// TIA Portal V19 export
// export: Created 2026-10-15T09:44:24.5896701Z, ExportSetting WithDefaults, DisplayName Totally Integrated Automation Portal, DisplayVersion V19, DisplayName TIA Portal Openness, DisplayVersion V19, DisplayName TIA Portal Version Control Interface, DisplayVersion V19, DisplayName STEP 7 Professional, DisplayVersion V19, DisplayName STEP 7 Safety, DisplayVersion V19, DisplayName WinCC Basic/Comfort/Advanced, DisplayVersion V19, DisplayName WinCC Unified, DisplayVersion V19
FUNCTION "ROLL_PB19" : Void   // FC27, SCL
{ S7_Optimized_Access := 'TRUE' }
VERSION : 0.1
// stored: AutoNumber true, IsIECCheckEnabled false, SetENOAutomatically false, UDAEnableTagReadback false
   VAR_TEMP
      r : Bool;
      a1 : Word;
      a2 : Word;
      activeDataBlock : Int;
      comparisonResults : Array[0..0] of Bool;
   END_VAR
BEGIN

   #r := FALSE;
   #a1 := W#16#0000;
   #a2 := W#16#0000;
   #activeDataBlock := 0;
   // PB19, STEP 5 network 1
   #r := ((NOT "ROLL_IO".Input[3, 6]) AND (NOT "ROLL_State".M[5, 6]) AND (NOT "ROLL_State".M[6, 0]) AND (NOT "ROLL_State".M[6, 2]) AND ("ROLL_IO".Input[3, 1] OR "ROLL_State".M[31, 5]) AND "ROLL_IO".Input[5, 2] AND "ROLL_IO".Input[5, 4] AND "ROLL_State".M[4, 1]);
   "ROLL_State".M[82, 0] := #r;
   // PB19, STEP 5 network 2
   #r := ((NOT "ROLL_IO".Input[3, 6]) AND (NOT "ROLL_State".M[12, 0]) AND (NOT "ROLL_State".M[5, 3]) AND (NOT "ROLL_State".M[5, 6]) AND ("ROLL_IO".Input[3, 1] OR "ROLL_State".M[31, 5]) AND "ROLL_IO".Input[8, 3] AND "ROLL_IO".Input[8, 5] AND "ROLL_State".M[4, 1]);
   "ROLL_State".M[82, 2] := #r;
   // PB19, STEP 5 network 3
   #r := ("ROLL_State".M[31, 5] AND "ROLL_State".M[40, 0]);
   IF #r THEN
       "ROLL_State".M[82, 3] := TRUE;
   END_IF;
   #r := (NOT "ROLL_State".M[31, 5]);
   IF #r THEN
       "ROLL_State".M[82, 3] := FALSE;
   END_IF;
   // PB19, STEP 5 network 4
   #r := ((NOT "ROLL_State".M[110, 1]) AND (NOT "ROLL_State".M[110, 2]) AND "ROLL_State".M[110, 0] AND "ROLL_State".M[110, 3] AND "ROLL_State".M[40, 0]);
   "ROLL_State".M[240, 0] := #r;
   // PB19, STEP 5 network 5
   #r := (((NOT "ROLL_State".M[110, 2]) AND "ROLL_State".M[110, 0] AND "ROLL_State".M[110, 1] AND "ROLL_State".M[110, 3] AND "ROLL_State".M[41, 1]) OR "ROLL_State".M[240, 0]);
   "ROLL_State".M[240, 0] := #r;
   // PB19, STEP 5 network 6
   #r := (((NOT "ROLL_State".M[110, 1]) AND "ROLL_State".M[110, 0] AND "ROLL_State".M[110, 2] AND "ROLL_State".M[110, 3] AND "ROLL_State".M[41, 1]) OR "ROLL_State".M[240, 0]);
   "ROLL_State".M[240, 0] := #r;
   // PB19, STEP 5 network 7
   #r := (("ROLL_State".M[110, 0] AND "ROLL_State".M[110, 1] AND "ROLL_State".M[110, 2] AND "ROLL_State".M[110, 3] AND "ROLL_State".M[41, 1]) OR "ROLL_State".M[240, 0]);
   "ROLL_State".M[240, 0] := #r;
   // PB19, STEP 5 network 8
   #r := ("ROLL_State".M[240, 0] AND "ROLL_State".M[31, 5]);
   IF #r THEN
       "ROLL_State".M[82, 4] := TRUE;
   END_IF;
   #r := ((NOT "ROLL_State".M[31, 5]) OR "ROLL_State".M[45, 5]);
   IF #r THEN
       "ROLL_State".M[82, 4] := FALSE;
   END_IF;
   // PB19, STEP 5 network 9
   #r := ((NOT "ROLL_IO".Output[17, 3]) AND (NOT "ROLL_State".M[82, 4]) AND (NOT "ROLL_State".S5Timers[91].Q) AND ("ROLL_State".M[82, 3] OR "ROLL_State".S5Timers[22].Q) AND "ROLL_IO".Input[8, 5]);
   "ROLL_IO".Output[17, 2] := #r;
   // PB19, STEP 5 network 10
   #r := ((NOT "ROLL_IO".Output[17, 2]) AND (NOT "ROLL_State".S5Timers[90].Q) AND "ROLL_IO".Input[3, 0] AND "ROLL_IO".Input[8, 5] AND "ROLL_State".M[82, 4]);
   "ROLL_IO".Output[17, 3] := #r;
   // PB19, STEP 5 network 11
   #a2 := #a1;
   #a1 := W#16#3060;
   #r := "ROLL_IO".Output[18, 0];
   "ROLL_TimerOp"(Number := 22,
                  Operation := 1,
                  Signal := #r,
                  Preset := #a1);
   // PB19, STEP 5 network 12
   #a2 := #a1;
   #a1 := W#16#1005;
   #r := "ROLL_IO".Output[17, 2];
   "ROLL_TimerOp"(Number := 90,
                  Operation := 1,
                  Signal := #r,
                  Preset := #a1);
   // PB19, STEP 5 network 13
   #a2 := #a1;
   #a1 := W#16#1040;
   #r := "ROLL_IO".Output[17, 3];
   "ROLL_TimerOp"(Number := 91,
                  Operation := 1,
                  Signal := #r,
                  Preset := #a1);
   // PB19, STEP 5 network 14
   #r := ((NOT "ROLL_State".M[12, 0]) AND (NOT "ROLL_State".M[19, 7]) AND ("ROLL_IO".Output[17, 2] OR "ROLL_IO".Output[17, 3] OR "ROLL_State".S5Timers[90].Q OR "ROLL_State".S5Timers[91].Q) AND ("ROLL_State".M[82, 3] OR "ROLL_State".M[82, 4]) AND "ROLL_IO".Input[8, 3] AND "ROLL_IO".Input[8, 4] AND "ROLL_State".M[82, 2]);
   "ROLL_IO".Output[18, 0] := #r;
   // PB19, STEP 5 network 15
   #r := "ROLL_IO".Output[18, 0];
   "ROLL_IO".Output[18, 1] := #r;
   // PB19, STEP 5 network 16
   #r := ("ROLL_IO".Output[18, 0] AND "ROLL_State".M[82, 4]);
   "ROLL_IO".Output[18, 2] := #r;
   // PB19, STEP 5 network 17
   #r := ("ROLL_IO".Output[18, 0] AND "ROLL_State".M[82, 4]);
   "ROLL_IO".Output[18, 3] := #r;
   // PB19, STEP 5 network 18
   RETURN;
END_FUNCTION
